# EPICS substitutions: iocs/motor/oms-asyn-ioc/db/MAXnet.substitutions
# C's iocOmsAsyn MAXnet.substitutions, P and PORT from st.cmd. C's PORT is
# MAXNET, the octet port, where devMotorAsyn finds no asynInt32 and the
# record fails init; PORT here is the omsMAXnetConfig port.
file "$(MOTOR)/db/asyn_motor.db"
{
pattern
{N,  M,       DTYP,         ADDR,  DESC,          EGU,  DIR,  VELO,  VBAS,  ACCL,  BDST,  BVEL,  BACC,  MRES,  PREC,  DHLM,  DLLM,  INIT}
{2,  "m$(N)", "asynMotor",  0,     "motor $(N)",  deg,  Pos,  10,    0,     .2,    0,     1,     2,     0.01,  5,     0,     0,     ""}
}
